FUNCTION_BLOCK ReliabilityIhm (* Reliability para a IHM: valor padrao ate chegar o primeiro valor do analisador *)
  (* Standard: 61499-2 *)
  (* Version 1.0, 05/11/2026, Hidryco, Hidryco, 1.0: Saida comeca em 80 (sensor sem MEASUREMENT IND. no SC1000, como pH e ORP, continua com 80); cada REQ copia Entrada para Saida e emite CNF. *)
  PACKAGE SE.Nereda;
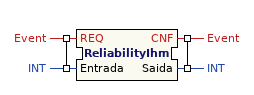
  EVENT_INPUT
    REQ WITH Entrada; (* Chegou valor de Reliability *)
  END_EVENT
  EVENT_OUTPUT
    CNF WITH Saida; (* Valor atualizado *)
  END_EVENT
  VAR_INPUT
    Entrada : INT; (* Reliability lido (MEASUREMENT IND.) *)
  END_VAR
  VAR_OUTPUT
    Saida : INT := 80; (* Reliability para a IHM *)
  END_VAR
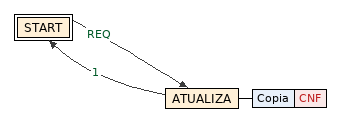
  EC_STATES
    START; (* Estado inicial *)
    ATUALIZA : Copia -> CNF; (* Copia o valor *)
  END_STATES
  EC_TRANSITIONS
    START TO ATUALIZA := REQ;
    ATUALIZA TO START := 1;
  END_TRANSITIONS
  ALGORITHM Copia IN ST: (* Saida := Entrada *)
Saida := Entrada;
  END_ALGORITHM
END_FUNCTION_BLOCK
